PROGRAM main
  VAR
    start AT %MX0.0 : BOOL;
    stop AT %MX0.1 : BOOL;
    prox AT %MX0.2 : BOOL;
    level AT %MX0.3 : BOOL;
    motor AT %QX0.0 : BOOL;
    solenoid AT %QX0.1 : BOOL;
    run_light AT %QX0.2 : BOOL;
    release : BOOL;
    mode_a AT %MX0.4 : BOOL;
    mode_b AT %MX0.5 : BOOL;
    mode_c AT %MX0.6 : BOOL;
    fill_light AT %QX0.3 : BOOL;
    full_light AT %QX0.4 : BOOL;
  END_VAR

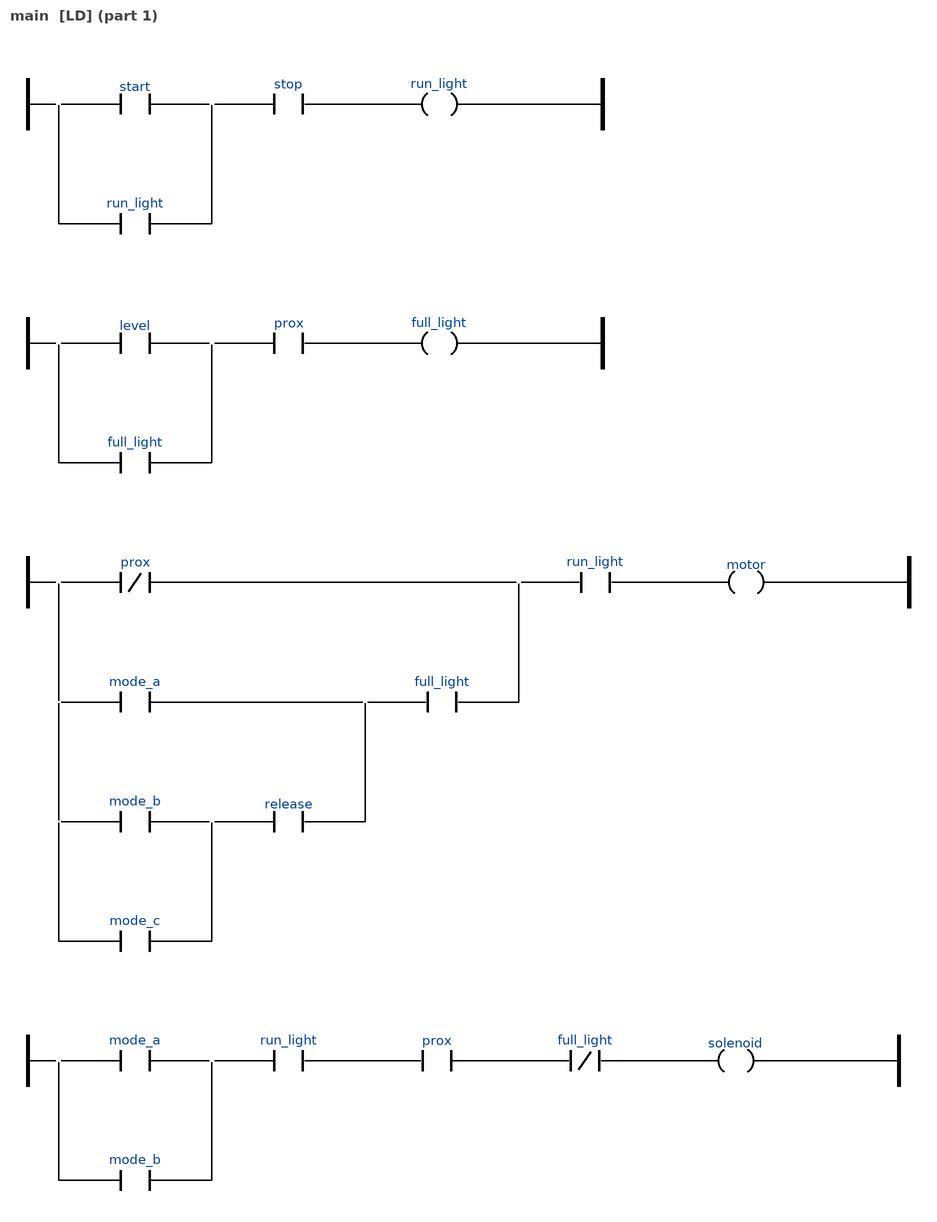
(* LD diagram, written out as Structured Text *)
run_light := (start OR run_light) AND stop;
full_light := (level OR full_light) AND prox;
motor := (NOT prox OR (mode_a OR (mode_b OR mode_c) AND release) AND full_light) AND run_light;
solenoid := (mode_a OR mode_b) AND run_light AND prox AND NOT full_light;
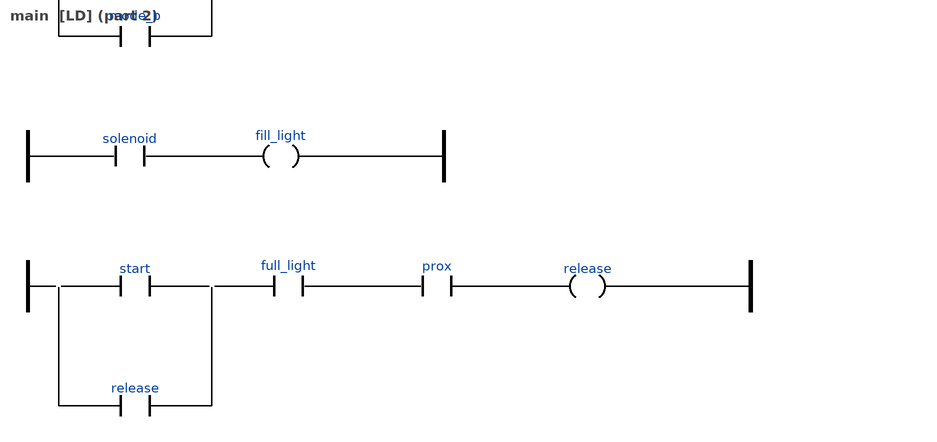
fill_light := solenoid;
release := (start OR release) AND full_light AND prox;
END_PROGRAM
